// Mitsubishi GX Works2 project: Practica f   PLC: FX3G

PROGRAM MAIN
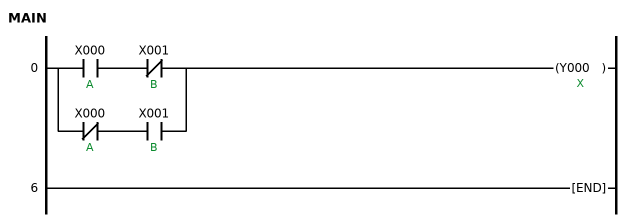
0     LD      X000  ; A
      ANI     X001  ; B
      LDI     X000  ; A
      AND     X001  ; B
      ORB
      OUT     Y000  ; X
6     END
END_PROGRAM
